TYPE ST_ParsedSignal :
STRUCT
    area                : E_MBArea;
    baseAddress         : UINT;
    bitIndex            : BYTE;
    registerCount       : UINT;
    dataType            : E_MBDataType;
    valid               : BOOL;
    isBitInRegister     : BOOL;
END_STRUCT
END_TYPE

(* stored: Version 1.1.0.1, ProductVersion 3.1.4024.0
   DUT ST_ParsedSignal: Id {569ede87-c53e-4b5c-b182-8e9e282ae5d2} *)
